Staubli VAL3: HMI_setting.pjx

--- HMI_setting.pjx ---
Parameters version=s8.15.3Cs9_BS3337 stackSize=5000 millimeterUnit=true
Program file=bind.pgx
Program file=main.pgx
Program file=moveTohome.pgx
Program file=onStart.pgx
Program file=seMaxJntForce.pgx
Program file=start.pgx
Program file=stop.pgx
Program file=teachHome.pgx
Program file=unLock.pgx
Data file=HMI_setting.dtx
Library alias=savedata path=Disk://source/saveData/saveData.pjx
Library alias=util path=Disk://HMI_cs9/HMI_util/HMI_util.pjx
Library alias=simulate path=Disk://HMI_cs9/simulate/simulate.pjx
Library alias=prog path=Disk://source/projectSource/program/program.pjx
Library alias=trajectory path=Disk://source/projectSource/trajectory/trajectory.pjx
Library alias=libTqe path=Disk://LibTorque/LibTorque.pjx
Library alias=rs path=Disk://source/projectSource/robotStatus/robotStatus.pjx

--- HMI_setting.dtx ---
mdesc mNomSpeed
bool bBack
bool bMove
bool bTeach
bool bSetup
string sLsit
string sSelTool
string sLastTool
string sList
string sUsingLib
string sLibList
bool bChangeLib
public bool bIsDoing
bool bToSave
bool bLock
bool bDisable[6]
bool bSetMaxJntForce
bool bSix_Axis
string sArmType
num nMaxJntForec[6]
string sArmDetail
string sPassword = "staubli2025"
string sBtnUnLock

--- main.pgx ---
public program main()
  local bool l_bExit
  local bool l_bResult
  local num l_nTool
  local tool l_tTool
  local num l_nUsingLib
  local num l_nResult
  local string l_sLib
  local num i
begin
  do
    if util:sPage!="setting"
      util:sPage="setting"
      call util:loadingPage()
      call onStart()
      call bind()
      userPage("setting")
      delay(0.5)
    endIf

    if sSelTool != sLastTool
      sLastTool=sSelTool
      toNum(sLastTool,l_nTool,l_bResult)
    endIf
    if bTeach
      bTeach=false
      call teachHome()
    elseIf bMove
      bMove=false
      call moveTohome()
    elseIf bSetup
      bSetup=false
      if l_nTool!=savedata:nJogTool
        savedata:nJogTool=l_nTool
        call savedata:setBaseJOG(l_nTool)
        savedata:libSave()
        delay(0.1)
      endIf
    elseIf bChangeLib
      bChangeLib=false
      if workingMode()!=1
        popUpMsg("请先将工作模式切换到手动模式")
      else
        l_sLib=delete(sUsingLib,3,0)
        toNum(l_sLib,l_nUsingLib,l_bResult)
        if !l_bResult
          return
        else
          bIsDoing=true
          savedata:nLibIndex=l_nUsingLib
          savedata:libSave()

          bToSave=true
          call prog:onSave(bToSave)
          bToSave=true
          call trajectory:onSave(bToSave)
          logMsg("手动开始切换:"+toString(".2",clock()))
          call prog:loadPROG(l_nUsingLib,l_nResult)
          call trajectory:loadTRAJ(l_nUsingLib,l_nResult)

          bIsDoing=false
        endIf
      endIf
    elseIf bBack
      bBack=false
      l_bExit=true
    endIf

    call libTqe:refresh()
    //    if bLock==true
    //      sBtnUnLock="解锁"
    //    else
    //      sBtnUnLock="保存"
    //    endIf
    delay(0)
  until l_bExit==true
end

--- start.pgx ---
program start()
begin
end

--- applyLib.pgx ---
public program applyLib()
begin
  savedata:bLibApplied=!savedata:bLibApplied
  savedata:libSave()
  delay(0.5)

end

--- bind.pgx ---
program bind()
begin
  userPageBindClick("setting","btnback",bBack,true)
  userPageBindClick("setting","btn1",bTeach,true)
  userPageBindClick("setting","btn2",bMove,true)
  userPageBindClick("setting","btn3",bSetup,true)
  userPageBind("setting","cbx1","options",sList,size(sList),"r")
  userPageBind("setting","cbx1","value",sSelTool,1,"rw")
  userPageBind("setting","cbx1_Copy1","options",sLibList,size(sLibList),"r")
  userPageBind("setting","cbx1_Copy1","value",sUsingLib,1,"rw")
  userPageBindClick("setting","btn3_Copy1",bChangeLib,true)
end

--- moveTohome.pgx ---
program moveTohome()
begin
  call simulate:simulateHome()
end

--- onStart.pgx ---
program onStart()
  local num l_i
  local string l_sPath
  local num i
begin
  l_sPath="Disk://data/CustomerLib"
  libList(l_sPath,sLibList)

  resize(sList,1,size(savedata:tToolItem))

  bIsDoing=false
  for l_i = 0 to size(sList)-1
    sList[l_i]=toString("",l_i)+","+savedata:tToolItem[l_i].sName
  endFor

  sSelTool=toString("",savedata:nUsingTool)+","+savedata:tToolItem[savedata:nUsingTool].sName
  sLastTool=""
//  bLock=true
//  sBtnUnLock="解锁"
//  //获取机器人类型
//  call libTqe:_getArmType(sArmType,sArmDetail)
//  if sArmType=="4_Axis"
//    resize(bDisable,1,4)
//    resize(nMaxJntForec,1,4)
//    bSix_Axis=false
//  elseIf sArmType=="6_Axis"
//    resize(bDisable,1,6)
//    resize(nMaxJntForec,1,6)
//    bSix_Axis=true
//  endIf
//  //初始化扭矩设置解锁按钮
//  for i=0 to size(bDisable)-1
//    bDisable[i]=true
//  endFor
  //  call libTqe:_getSetForce(nMaxJntForec)
  call libTqe:initParameter()
end

--- seMaxJntForce.pgx ---
program seMaxJntForce()
  local num i
begin
//  if sArmType=="4_Axis"
//    for i=0 to 3
//      libTqe:tArm4Force[sArmDetail].nMaxJnt4Force[i]=nMaxJntForec[i]
//    endFor
//  elseIf sArmType=="6_Axis"
//    for i=0 to 5
//      libTqe:tArm6Force[sArmDetail].nMaxJnt6Force[i]=nMaxJntForec[i]
//    endFor
//  endIf
//  libTqe:libSave()
//  delay(0.1)
end

--- stop.pgx ---
program stop()
begin
end

--- teachHome.pgx ---
public program teachHome()
  local bool l_bResult
begin
  l_bResult=userPageConfirm("是否记录当前位置为home位置？")
  if l_bResult
    savedata:jHome=herej()
    savedata:libSave()
    delay(0.1)
    popUpMsg("home位置已记录并保存")
  endIf
end

--- unLock.pgx ---
program unLock()
  local string l_sEntry
  local bool l_bResult
  local num i
begin
//  if bLock==true
//    l_bResult=userPagePrompt("请输入密码",l_sEntry)
//    if l_bResult==false
//      return
//    endIf
//    if l_sEntry!=sPassword[0]
//      popUpMsg("密码错误")
//      return
//    endIf
//    //2024.04.29 add解锁扭矩限位设置
//    for i=0 to size(bDisable)-1
//      bDisable[i]=false
//    endFor
//    popUpMsg("修改后请点击保存!")
//    bLock=false
//  else
//    for i=0 to size(bDisable)-1
//      bDisable[i]=true
//    endFor
//    call seMaxJntForce()
//    call libTqe:_getSetForce(nMaxJntForec)
//    popUpMsg("机器人关节扭矩限制保存成功!")
//    bLock=true
//  endIf
end
